(* CODESYS project SysParSafety.xml

Project tree, tasks and I/O mapping:
  visualisation SysParSafety
*)

// /SysParSafety
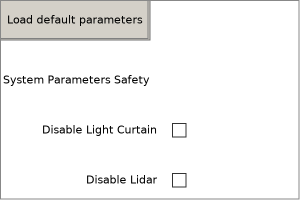
VISUALIZATION SysParSafety  // 300x200
    Button (0,0 150x40), "Load default parameters"
        tap PRG_VisuTask_10ms._fbParametersCtrl._btnLoadDefaultParameters.xbtn
    Label (0,60 300x40), "System Parameters Safety"
    Checkbox (170,110 40x40), variable: PersistentVars.scSafety.xDisableLightCurtains
    Label (10,110 150x40), "Disable Light Curtain"
    Label (10,160 150x40), "Disable Lidar"
    Checkbox (170,160 40x40), variable: PersistentVars.scSafety.xDisableLidar
END_VISUALIZATION
